(* IEC 61131-3 sources: 2026_Projet_YGO_ExcavatriceDragage/CODE/J_SUPERVISION/_TYPES/4_JOYSTICK_ACQUISITION, 16 files *)

(* ---- E_ArmingBlockReason.st ---- *)
(* =======================================================================
   🚦 E_ArmingBlockReason — Motif de blocage de l'armement joystick
   ───────────────────────────────────────────────────────────────
   🎯 Rôle : dire EN CLAIR pourquoi ArmingPermit est FALSE, pour l'IHM et
      le troubleshooting (« pourquoi je ne peux pas armer »).
   📄 Doc : DOC/AF/AF_Partie-08_Fonction_Joystick_v2.5.md §7
   ======================================================================= *)
TYPE E_ArmingBlockReason :
(
    NONE            := 0,   // Armement possible (au moins un axe x sens dispo)
    MODE_DISABLE    := 1,   // Mode DISABLE
    POWER_CUTOFF    := 2,   // Coupure puissance amont (M1/M2/M3)
    CONTACTOR_OFF   := 3,   // Chaîne AU non réarmée (PowerContactorEngaged FALSE)
    BUCKET_BUSY     := 4,   // Action benne en cours (+ 1 scan de fin d'action)
    ALL_AXES_BLOCKED := 5   // Base OK mais aucun axe x sens sélectionné n'est disponible
);
END_TYPE

(* ---- ST_AcquisitionEncoderQualified.st ---- *)
(* ═══════════════════════════════════════════════════════════════
   🧲 ST_AcquisitionEncoderQualified — Façade codeur qualifiée
   ───────────────────────────────────────────────────────────────
   🎯 Rôle : Encapsuler les mesures métriques, statuts de référencement,
      défauts et signaux hardware produits par FB_Encoder dans PRG_02_Acquisition.
   📤 Producteur unique : PRG_02_Acquisition (Data.EncoderM1 / Data.EncoderM2).
   📄 Doc : DOC/AF/AF_Partie-06_Acquisition_Qualification_IO_v2.4.md
   ═══════════════════════════════════════════════════════════════ *)

TYPE ST_AcquisitionEncoderQualified :
STRUCT
    Measurement              : ST_fbEncoder_Measurement; // 📊 Mesure métrique (CablePosM, SpeedMps, etc.)
    Ready                    : BOOL;                     // 🟢 Façade codeur prête
    Fault                    : ST_Fault;                 // ❌ Diagnostic défaut codeur
    Homed                    : BOOL;                     // 🎯 Codeur référencé
    HomingSuspect            : BOOL;                     // ⚠️ Référencement suspect
    EncoderFault             : BOOL;                     // ❌ Défaut fiabilité (indisponible ou incohérent)
    HomedAndReliable         : BOOL;                     // ✅ Référencé ET fiable (sans incohérence)
    PresetConfirmationFailed : BOOL;                     // ❌ Échec confirmation preset
    HwOut                    : ST_fbEncoder_HwOut;       // 📡 Commandes hardware de preset (lecture seule)
END_STRUCT
END_TYPE

(* ---- ST_AcquisitionInterPrg.st ---- *)
(* ═══════════════════════════════════════════════════════════════
   🧲 ST_AcquisitionInterPrg — Bus d'échange inter-PRG produit par PRG_02_Acquisition
   ───────────────────────────────────────────────────────────────
   🎯 Rôle : Encapsuler les mesures câbles/vitesses, les états joystick qualifiés,
      les positions M3 et les diagnostics DI publiés par PRG_02_Acquisition vers
      les consommateurs (PRG_03/04/05/07, FB_TroubleshootingView).
   📤 Producteur unique : PRG_02_Acquisition (VAR_OUTPUT Data : ST_AcquisitionInterPrg).
   📄 Doc : DOC/AF/AF_Partie-06_Acquisition_Qualification_IO_v2.4.md
   🔌 Architecture : Bus de données typé — encapsulation des échanges inter-PRG.
   ═══════════════════════════════════════════════════════════════ *)

TYPE ST_AcquisitionInterPrg :
STRUCT
    // === 🛡️ Drapeau de vie & validité globale des données ===
    DataValid                    : BOOL; // 🟢 TRUE = PRG_02 a complété son scan et les données sont fraîches et qualifiées

    // === 📦 Structures qualifiées du bus ===
    Joystick                     : ST_AcquisitionJoystickQualified;    // 🕹️ Données et commandes joystick qualifiées
    Network                      : ST_AcquisitionNetworkDiagnostics;  // 🔌 Diagnostics réseaux CANopen et EtherCAT
    EncoderM1                    : ST_AcquisitionEncoderQualified;     // 🧲 Façade codeur qualifiée M1 (Retenue)
    EncoderM2                    : ST_AcquisitionEncoderQualified;     // 🧲 Façade codeur qualifiée M2 (Benne)
    MachineHoming                : ST_MachineHoming;                   // 🎯 État homing conjoint machine (M1/M2/benne)

    // === 🩺 Diagnostics modules E/S ===
    InputModules                 : ST_IOModuleDiag; // 🩺 Diagnostic carte des 5 modules E/S (AF06 §3bis)

    // === 🧪 Simulation & variateur M3 filtré ===
    InputSource                  : ST_InputSource; // 🔀 Flags de bascule de source (réel/simu) par domaine
    M3                           : ST_M3DriveFeedback; // ↔️ Retours variateur M3 filtrés (consommé PRG_05)
END_STRUCT
END_TYPE

(* ---- ST_AcquisitionJoystickQualified.st ---- *)
(* ═══════════════════════════════════════════════════════════════
   🕹️ ST_AcquisitionJoystickQualified — Données joystick qualifiées
   ───────────────────────────────────────────────────────────────
   🎯 Rôle : Encapsuler les commandes d'axes, statut homme-mort et diagnostics
      produits par FB_Joystick dans PRG_02_Acquisition.
   📤 Producteur unique : PRG_02_Acquisition (Data.Joystick).
   📄 Doc : DOC/AF/AF_Partie-06_Acquisition_Qualification_IO_v2.4.md
   ═══════════════════════════════════════════════════════════════ *)

TYPE ST_AcquisitionJoystickQualified :
STRUCT
    AxisX               : ST_fbJoystick_AxisCmd; // 📊 Commande et direction qualifiée axe X
    AxisY               : ST_fbJoystick_AxisCmd; // 📊 Commande et direction qualifiée axe Y
    DeadmanArmed        : BOOL;                  // 🔒 Homme-mort armé et valide
    AtNeutralXY         : BOOL;                  // 🟢 Les deux axes X et Y sont au neutre
    ArmingPermitDenied  : BOOL;                  // ⚠️ Tentative d'armement sans permission
    Ready               : BOOL;                  // 🟢 Façade joystick prête et opérationnelle
    Fault               : ST_Fault;              // ❌ Diagnostic défaut joystick
    NeutralXAct         : INT;                   // 📍 Valeur ADC neutre calibré X
    NeutralYAct         : INT;                   // 📍 Valeur ADC neutre calibré Y
END_STRUCT
END_TYPE

(* ---- ST_AcquisitionNetworkDiagnostics.st ---- *)
(* ═══════════════════════════════════════════════════════════════
   🔌 ST_AcquisitionNetworkDiagnostics — Diagnostics réseaux qualifiés
   ───────────────────────────────────────────────────────────────
   🎯 Rôle : Encapsuler les états opérationnels et diagnostics des bus CANopen
      et EtherCAT produits par PRG_02_Acquisition.
   📤 Producteur unique : PRG_02_Acquisition (Data.Network).
   📄 Doc : DOC/AF/AF_Partie-06_Acquisition_Qualification_IO_v2.4.md
   ═══════════════════════════════════════════════════════════════ *)

TYPE ST_AcquisitionNetworkDiagnostics :
STRUCT
    CanOpenMaster   : ST_Diag_Device; // 🔌 Diagnostic maître CANopen
    Joystick        : ST_Diag_Device; // 🕹️ Diagnostic esclave Joystick MCB560
    EthercatMaster  : ST_Diag_Device; // 🔌 Diagnostic maître EtherCAT
    EncoderM1       : ST_Diag_Device; // 🧲 Diagnostic esclave Codeur M1 (COD1)
    EncoderM2       : ST_Diag_Device; // 🧲 Diagnostic esclave Codeur M2 (COD2)
    DriveM3         : ST_Diag_Device; // ⚙️ Diagnostic esclave Variateur M3 (AC600)
END_STRUCT
END_TYPE

(* ---- ST_ArmingAvailability.st ---- *)
(* =======================================================================
   🚦 ST_ArmingAvailability — Disponibilité de mouvement par axe et sens
   ───────────────────────────────────────────────────────────────
   🎯 Rôle : dire, pour chaque axe x sens, si le mouvement peut REELLEMENT
      partir (permis effectif + pas de SafeStop/faute de CET axe). Sert de
      base honnête à ArmingPermit (au moins un dispo) et de diagnostic
      « pourquoi ça bloque » pour l'IHM / le troubleshooting.
   📤 Producteur : PRG_04_Treuils_Benne (agrège M1/M2 + lit M3 via bus PRG_05, lag 1 scan).
   📄 Doc : DOC/AF/AF_Partie-08_Fonction_Joystick_v2.5.md §7
   ======================================================================= *)
TYPE ST_ArmingAvailability :
STRUCT
    M1AscentAvail      : BOOL;   // TRUE = montée M1 peut partir
    M1DescendAvail     : BOOL;   // TRUE = descente M1 peut partir
    M2AscentAvail      : BOOL;   // TRUE = montée/fermeture M2 peut partir
    M2DescendAvail     : BOOL;   // TRUE = descente/ouverture M2 peut partir
    M3TremieAvail      : BOOL;   // TRUE = translation M3 vers trémie peut partir
    M3MaintenanceAvail : BOOL;   // TRUE = translation M3 vers maintenance peut partir
    AnyAxisAvail       : BOOL;   // OR des 6 — au moins une action peut partir (condition d'armement)
    BlockedReason      : E_ArmingBlockReason;   // Motif si armement impossible
END_STRUCT
END_TYPE

(* ---- ST_EncoderHMI.st ---- *)
(* ═══════════════════════════════════════════════════════════════
   🧲 ST_EncoderHMI — Données d'échange IHM pour les codeurs absolus
   ───────────────────────────────────────────────────────────────
   🎨 Destiné à l'affichage des informations et diagnostics des codeurs.
   ═══════════════════════════════════════════════════════════════ *)
TYPE ST_EncoderHMI :
STRUCT
    RawPos           : UDINT; (* 📊 Position brute lue sur le bus *)
    Alarms           : UINT;  (* ⚠️ Code d'alarme brut du codeur *)
    Warnings         : UINT;  (* 🟧 Code d'avertissement brut du codeur *)
    SlaveOperational : BOOL;  (* 📡 Esclave EtherCAT opérationnel *)
    PresetTriggerCmd : WORD;  (* 🎯 Commande de preset active *)
    PresetValueOut   : UDINT; (* 📐 Valeur de preset envoyée au codeur *)
    Error            : BOOL;  (* Codeur en défaut (liaison EtherCAT ou preset) *)
    ErrorId          : WORD;  (* ❌ Code défaut codeur *)

    (* 🎯 Homing — prise d'origine / référencement *)
    Homed                   : BOOL;             (* 🎯 Prise d'origine (Homing) validée *)
    HomingBusy              : BOOL;             (* ⏳ Référencement en cours *)
    HomingDone              : BOOL;             (* ✅ Pulse de référencement réussi *)
    HomingError             : BOOL;             (* Défaut de référencement *)
    HomingErrorId           : WORD;             (* ❌ Bitfield défaut homing *)
    HomingState             : E_State;          (* 🤖 État FB_Encoder_Homing *)
    HomingStateAtError      : E_State;          (* 🧭 État lors du défaut *)
    HomingSuspect           : BOOL;             (* ⚠️ Référence à confirmer *)
    HomingRefRaw            : UDINT;            (* 📐 Référence brute appliquée *)
END_STRUCT
END_TYPE

(* ---- ST_HardwareImage.st ---- *)
(* ═══════════════════════════════════════════════════════════════
   🏗️ ST_HardwareImage — Structure globale d'image matérielle (Frontière HwIn)
   ───────────────────────────────────────────────────────────────
   🎨 Agrège les 4 sous-domaines matériels : Winch, Translation, Operator, Machine.
   ═══════════════════════════════════════════════════════════════ *)
TYPE ST_HardwareImage :
STRUCT
    Winch       : ST_HwWinch;       (* Entrées brutes domaine Treuils M1/M2 + codeurs *)
    Translation : ST_HwTranslation; (* Entrées brutes domaine Translation M3 + variateur *)
    Operator    : ST_HwOperator;    (* Entrées brutes domaine Opérateur / Joystick / bus CAN *)
    Machine     : ST_HwMachine;     (* Entrées brutes domaine Sécurités/Communs Machine *)
END_STRUCT
END_TYPE

(* ---- ST_HwMachine.st ---- *)
(* ═══════════════════════════════════════════════════════════════
   🏗️ ST_HwMachine — Image matérielle brute des entrées communes Machine
   ───────────────────────────────────────────────────────────────
   🎨 Regroupe les signaux physiques d'entrée bruts communs à la machine.
   ═══════════════════════════════════════════════════════════════ *)
TYPE ST_HwMachine :
STRUCT
    PowerContactorEngaged_DI       : BOOL; (* Confirm. contacteur puissance engagé *)
    EmergencyChainClosed_DI        : BOOL; (* Boucle AU fermée (coup-de-poing + contact PLC) *)
    PhaseRotationOk_DI             : BOOL; (* Contrôle rotation phases élec. OK *)
    M1_M2_M3_BrakeThermalOk_DI     : BOOL; (* Thermique frein M1/M2/M3 commun OK *)
    M1_M2_KoboldBottomTouch_DI     : BOOL; (* Retour détecteur fond Kobold *)
    HydraulicThermalOk_DI          : BOOL; (* Thermique centrale hydraulique OK *)
    ConveyorInfeedReady_DI         : BOOL; (* Autorisation démarrage crible (dépôt gravats) *)
    TremieFull_OR_GateRaised_DI    : BOOL; (* : Trémie pleine OU grille levée — pas encore câblé électriquement,
                                               déclaré en avance (Device_IO_20260826). Aucun consommateur pour l'instant :
                                               l'interdiction translation M3→Trémie est une tâche à part, voir PLAN_TASK.md. *)
END_STRUCT
END_TYPE

(* ---- ST_HwOperator.st ---- *)
(* ═══════════════════════════════════════════════════════════════
   🏗️ ST_HwOperator — Image matérielle brute des entrées Opérateur / Joystick
   ───────────────────────────────────────────────────────────────
   🎨 Regroupe les signaux physiques d'entrée bruts du joystick CANopen JOY1.
   ═══════════════════════════════════════════════════════════════ *)
TYPE ST_HwOperator :
STRUCT
    JoyXRaw_ANA1      : INT;          (* Valeur brute analogique axe X (Translation) *)
    JoyYRaw_ANA2      : INT;          (* Valeur brute analogique axe Y (Levage) *)
    JoyBtnRaw         : BOOL;         (* Bouton brut joystick (Homme-Mort) *)
    CanBusState       : INT;          (* État bus CANopen (CANbus.GetBusState) *)
    JOY1_DeviceState  : DEVICE_STATE; (* État device JOY1 (GetDeviceState) *)
END_STRUCT
END_TYPE

(* ---- ST_InputSource.st ---- *)
(* ═══════════════════════════════════════════════════════════════
   🔀 ST_InputSource — Flags de bascule de source (réel/simu) par domaine
   ───────────────────────────────────────────────────────────────
   🎯 Rôle : Regrouper les 4 impulsions 1 cycle signalant qu'une source
      d'entrée a basculé (réel ↔ simu) pour un domaine donné.
   📤 Producteur unique : PRG_02_Acquisition (Data.InputSource).
   📥 Consommateur : PRG_07_Supervision (Data.InputSource.* → GVL_IHM).
   📄 Doc : DOC/AF/AF_Partie-06_Acquisition_Qualification_IO_v2.4.md
   🔌 Architecture : Bus de données typé — encapsulation des échanges inter-PRG.
   ═══════════════════════════════════════════════════════════════ *)

TYPE ST_InputSource :
STRUCT
    WinchInputSourceChanged       : BOOL; // 🔀 Source Winch a basculé (réel/simu)
    TranslationInputSourceChanged: BOOL; // 🔀 Source Translation a basculé
    OperatorInputSourceChanged   : BOOL; // 🔀 Source Opérateur a basculé
    MachineInputSourceChanged    : BOOL; // 🔀 Source Machine a basculé
END_STRUCT
END_TYPE

(* ---- ST_JoystickChecklist.st ---- *)
(* ═══════════════════════════════════════════════════════════════
   🕹️ ST_JoystickChecklist — Diagnostic chronologique communication & prise en main Joystick
   ───────────────────────────────────────────────────────────────
   🎨 Permet de vérifier la chaîne Joystick (CANopen, Homme-mort, Neutre, Calibration).
   ═══════════════════════════════════════════════════════════════ *)
TYPE ST_JoystickChecklist :
STRUCT
    (* 1. Bus & Matériel *)
    Step1_CanBusActive           : BOOL; (* TRUE = Bus CANopen en état ACTIVE *)
    Step2_JoystickOperational    : BOOL; (* TRUE = Esclave JOY1 en état RUNNING *)

    (* 1bis. Entrées physiques directes HwIn *)
    HwIn_JoyBtnRaw_DI            : BOOL; (* Bouton brut homme-mort issu de HwIn.Operator *)
    NeutralXAct                  : BOOL; (* TRUE = Axe X au neutre (PRG_02_Acquisition.Data.Joystick.AxisX.Direction = 0) *)
    NeutralYAct                  : BOOL; (* TRUE = Axe Y au neutre (PRG_02_Acquisition.Data.Joystick.AxisY.Direction = 0) *)

    (* 2. Prise en main & Sécurité *)
    Step3_DeadmanPressed         : BOOL; (* TRUE = Bouton Homme-Mort appuyé *)
    Step4_NeutralAcquired        : BOOL; (* TRUE = Repassé par le neutre (autorisation mouvement) *)
    DeadmanArmed                 : BOOL; (* TRUE = Homme-Mort armé avec passage au neutre validé *)

    (* 3. Éligibilité globale *)
    AllConditionsMet             : BOOL; (* TRUE = Joystick prêt pour piloter un axe *)
    JoystickSelected             : BOOL; (* TRUE = Joystick maître sélectionné IHM *)
    SelJoystickWinch             : INT;  (* Sélection Treuil (0=Couplé M1+M2, 1=M1 seul, 2=M2 seul) *)

    (* 4. Mesures brutes & Filtrées *)
    RawX                         : INT;  (* Valeur brute axe X (0..10000) *)
    RawY                         : INT;  (* Valeur brute axe Y (0..10000) *)
    DeflectionX_Pct              : REAL; (* Déflexion signée X (%) *)
    DeflectionY_Pct              : REAL; (* Déflexion signée Y (%) *)
    DirectionX                   : INT;  (* Direction filtrée X (-1 / 0 / +1) *)
    DirectionY                   : INT;  (* Direction filtrée Y (-1 / 0 / +1) *)
END_STRUCT
END_TYPE

(* ---- ST_JoystickCmd.st ---- *)
(* ═══════════════════════════════════════════════════════════════
   🎮 ST_JoystickCmd — Commandes IHM pour le Joystick
   ═══════════════════════════════════════════════════════════════ *)
TYPE ST_JoystickCmd :
STRUCT
    Calibrate : BOOL; (* 🎯 Demande de recalage au neutre (front) *)
END_STRUCT
END_TYPE

(* ---- ST_JoystickHMI.st ---- *)
(* ═══════════════════════════════════════════════════════════════
   🕹️ ST_JoystickHMI — Données d'échange IHM pour le Joystick
   ───────────────────────────────────────────────────────────────
   📄 Structuration en Cmd / State / Cfg , homogène avec ST_ModesHMI.
   Cfg = réglages FB_Joystick éditables IHM (deadband, temporisations), pontés vers
   GVL_PERSISTENT via FB_CfgPersistBridge_fbJoystick_Cfg. La calibration du neutre reste
   dans GVL_PERSISTENT (bouton Calibrate). Pas de Bypass (concept absent de ce struct).
   ═══════════════════════════════════════════════════════════════ *)
TYPE ST_JoystickHMI :
STRUCT
    Cmd   : ST_JoystickCmd;
    State : ST_JoystickState;
    Cfg   : ST_fbJoystick_Cfg;
END_STRUCT
END_TYPE

(* ---- ST_JoystickState.st ---- *)
(* ═══════════════════════════════════════════════════════════════
   🚦 ST_JoystickState — États et diagnostics IHM du Joystick
   ═══════════════════════════════════════════════════════════════ *)
TYPE ST_JoystickState :
STRUCT
    RawX         : INT;        (* 🕹️ Axe X brut du joystick (0..10000) *)
    RawY         : INT;        (* 🕹️ Axe Y brut du joystick (0..10000) *)
    RawButton    : BOOL;       (* 🔘 Bouton homme-mort brut *)
    AxisCmdX     : ST_fbJoystick_AxisCmd; (* ⚙️ Consigne d'axe X normalisée (sortie FB_Joystick) *)
    AxisCmdY     : ST_fbJoystick_AxisCmd; (* ⚙️ Consigne d'axe Y normalisée (sortie FB_Joystick) *)
    NeutralXAct  : INT;        (* 🎯 Neutre X calibré actuel (lecture seule) *)
    NeutralYAct  : INT;        (* 🎯 Neutre Y calibré actuel (lecture seule) *)
    DeadmanArmed : BOOL;       (* 🔫 Geste homme-mort armé (FB_Joystick.DeadmanArmed) *)
    AtNeutral    : BOOL;       (* : TRUE si les 2 axes sont en zone morte (position centrale) *)
    Online       : BOOL;       (* 📡 Liaison CAN joystick active *)
    Operational  : BOOL;       (* 🟢 Joystick opérationnel *)
    Error        : BOOL;       (* Joystick en défaut *)
    ErrorId      : WORD;       (* ❌ Code défaut joystick *)
END_STRUCT
END_TYPE

(* ---- ST_M3DriveFeedback.st ---- *)
(* ═══════════════════════════════════════════════════════════════
   ↔️ ST_M3DriveFeedback — Retours variateur M3 filtrés
   ───────────────────────────────────────────────────────────────
   🎯 Rôle : Encapsuler les retours variateur M3 (mot d'état + fréquence réelle)
      conditionnés par PRG_02_Acquisition et consommés par PRG_05_Translation.
   📤 Producteur unique : PRG_02_Acquisition (Data.M3).
   📥 Consommateur : PRG_05_Translation (Data.M3.StatusWord / Data.M3.ActualFrequencyHz).
   📄 Doc : DOC/AF/AF_Partie-06_Acquisition_Qualification_IO_v2.4.md
   🔌 Architecture : Bus de données typé — encapsulation des échanges inter-PRG.
   ═══════════════════════════════════════════════════════════════ *)

TYPE ST_M3DriveFeedback :
STRUCT
    StatusWord        : UINT; // 📊 Mot d'état variateur M3 filtré
    ActualFrequencyHz : UINT; // 📊 Fréquence réelle M3 filtrée
END_STRUCT
END_TYPE
